INTERFACE I_EquipmentModule EXTENDS I_Diagnosable

METHOD StartCycle                   // one cycle; taken up as soon as the module is ready
END_METHOD

PROPERTY IsCycleDone : BOOL
GET
END_GET
END_PROPERTY

END_INTERFACE

(* stored: Version 1.1.0.1
   Itf I_EquipmentModule: Id {c6aedb48-414c-4e59-8fef-f768cb1b1042}
   Method StartCycle: Id {2f89702c-ce7a-47fd-801e-26186d5610c4}
   Property IsCycleDone: Id {4bdf95de-2ceb-4496-9123-08730d61480e}
   Get Get: Id {8f52e5b5-374b-4cf5-b76a-7a6dcb4d78df} *)
